FUNCTION_BLOCK EEE_Bruto (* Elevatoria de esgoto bruto - HidrycoLib *)
  (* Standard: 61499-2 *)
  (* Version 1.9, 21/10/2026, Hidryco, Hidryco, 1.9: Necessidade recebe o nivel em % (STS_NIVEL) para o grafico das faixas. 1.8: PID de nivel e velocidades da IHM/SCADA em Hz (conversao no CLP). 1.7: faixas da Necessidade e PID de nivel em % da altura do poco (LIT_100_03.stsPorcentagem). 1.6: pidCtl PidNivel com CycleTime 1000 ms (sem ele o calculo ciclico do pidSC ficava sem periodo). 1.5: variaveis de controle nos sub-CATs Necessidade, Revezamento e PID (padrao ElevatoriaEsgotoBruto); reset cmdResetFalhas / E_RESET_FALHAS_PROCESSO; PT_100_01, LSL_100_04, LSH_100_05 e pidCtl PidNivel. 1.4: simbolos sBoiaL/sBoiaH (boias animadas, verde/vermelho); velocidades na IHM em Hz. 1.3: selecao do gerador bomba por bomba (geradorHabilitaBS01/02/03, cada uma so na sua bomba; antes geradorHabilita unica). 1.2: emergencia do PCM NF (stsEmergenciaPainel FALSE = em emergencia, so depois da 1a leitura); FALHA UCP das bombas NF (cfgTermicaNF TRUE: FALSE no campo = falha); rede do CAT reorganizada. 1.1: emergencia do PCM pelo symlink ${PATH}stsEmergenciaPainel (soma com stsEmergencia do processo); comunicacao dos ATV630 pelos symlinks ${PATH}atvComunicacaoBS01..03 (ComStatus do HW CAT ATVSpeedControlMbtcp) publicada como ${PATH}BS_100_0x.stsFalhaComunicacao; cfgUsaFalhaComunicacao TRUE; estado 7 = emergencia. 1.0: elevatoria de esgoto bruto (3 bombas 100-BS-01/02/03, 2 + 1 reserva). Faixas de nivel do LIT-03, revezamento por tempo, velocidade pelo PID de nivel, HH do Nereda segura o esgoto ate o H do poco, operacao pelas boias com o LIT-03 em falha, falha de recalque pelo PIT-01. Campo por symlink ${PATH}: stsBoiaNivelBaixo (LSL-04), stsBoiaNivelAlto (LSH-05); bombas e sensores pelos symlinks dos proprios CATs (${PATH}BS_100_0x., ${PATH}LIT_100_03., ${PATH}PIT_100_01.). *)
  PACKAGE Hidryco.HidrycoLib;
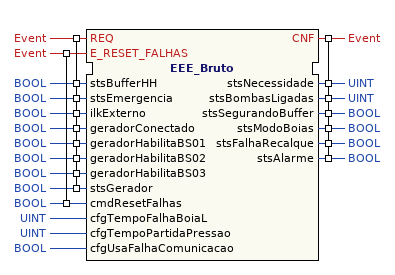
  EVENT_INPUT
    REQ WITH stsBufferHH, stsEmergencia, ilkExterno, geradorConectado, geradorHabilitaBS01, geradorHabilitaBS02, geradorHabilitaBS03, stsGerador; (* Atualizacao do processo *)
    E_RESET_FALHAS WITH cmdResetFalhas; (* Reset pelo processo (elevatoria, bombas e sensores) com cmdResetFalhas = TRUE *)
  END_EVENT
  EVENT_OUTPUT
    CNF WITH stsNecessidade, stsBombasLigadas, stsSegurandoBuffer, stsModoBoias, stsFalhaRecalque, stsAlarme; (* Status (so na mudanca) *)
  END_EVENT
  VAR_INPUT
    stsBufferHH : BOOL; (* Alarme HH do nivel do tanque de equalizacao do Nereda (40-LT-0001): a elevatoria segura o esgoto *)
    stsEmergencia : BOOL; (* Emergencia pelo processo (soma com a emergencia do PCM lida pelo symlink stsEmergenciaPainel): retira o comando das bombas *)
    ilkExterno : BOOL; (* Intertravamento externo do automatico das bombas (ex.: falha das UCTs, futuro) *)
    geradorConectado : BOOL; (* O gerador pode alimentar as bombas *)
    geradorHabilitaBS01 : BOOL; (* Bomba 100-BS-01 liberada para operar com a planta no gerador (HAB_BS_100_01 do CAT Subestacao) *)
    geradorHabilitaBS02 : BOOL; (* Bomba 100-BS-02 liberada para operar com a planta no gerador (HAB_BS_100_02 do CAT Subestacao) *)
    geradorHabilitaBS03 : BOOL; (* Bomba 100-BS-03 liberada para operar com a planta no gerador (HAB_BS_100_03 do CAT Subestacao) *)
    stsGerador : BOOL; (* Planta alimentada pelo gerador *)
    cmdResetFalhas : BOOL; (* TRUE = reset (com o evento E_RESET_FALHAS) *)
    cfgTempoFalhaBoiaL : UINT := 10; (* Operacao pelas boias com a boia LSL com defeito: bombas ficam ligadas este tempo (min) depois que a LSH desce *)
    cfgTempoPartidaPressao : UINT := 30; (* Alarmes L/LL do PIT-01 inibidos ate a bomba estar ligada ha este tempo (s); tambem inibidos com as bombas paradas *)
    cfgUsaFalhaComunicacao : BOOL := TRUE; (* Bombas: TRUE = falha de comunicacao com o ATV630 (symlink atvComunicacaoBS0x = ComStatus do HW CAT) tira a bomba do automatico *)
  END_VAR
  VAR_OUTPUT
    stsNecessidade : UINT; (* Numero de bombas pedidas (0, 1, 2) *)
    stsBombasLigadas : UINT; (* Bombas ligadas *)
    stsSegurandoBuffer : BOOL; (* Elevatoria parada segurando o esgoto (HH do tanque do Nereda) *)
    stsModoBoias : BOOL; (* Operacao de emergencia pelas boias (LIT-03 em falha) *)
    stsFalhaRecalque : BOOL; (* Falha de recalque (pressao LL com bomba ligada) - memorizada ate o reset *)
    stsAlarme : BOOL; (* Algum alarme da elevatoria *)
  END_VAR
  FBS
    IThis : EEE_Bruto_HMI(QI := TRUE);
    plcStart1 : plcStart(Prio := 10);
    Logica : basicEEEBruto;
    Tick : E_CYCLE(DT := T#1s);
    PidNivel : pidCtl(CycleTime := 1000, Direction := FALSE, Bump := FALSE, ProhibitOutInc := FALSE, ProhibitOutDec := FALSE);
    LIT_100_03 : Sensor_Generico(pin_FC98F78ABCBC0A7E := TRUE, pin_CC8EEC06FF0C4430 := 'm');
    PT_100_01 : Sensor_Generico(pin_CC8EEC06FF0C4430 := 'bar');
    LSL_100_04 : SYMLINKMULTIVARDST_1559B0FF8170C9BA0(NAME1 := '$${PATH}stsBoiaNivelBaixo', QI := TRUE); {SET_ATTRIBUTE(Configuration.GenericFBType.InterfaceParams, Runtime.System#I:=1;VALUE${I$}:BOOL)}
    LSH_100_05 : SYMLINKMULTIVARDST_1559B0FF8170C9BA0(NAME1 := '$${PATH}stsBoiaNivelAlto', QI := TRUE); {SET_ATTRIBUTE(Configuration.GenericFBType.InterfaceParams, Runtime.System#I:=1;VALUE${I$}:BOOL)}
    EmergenciaPainel : SYMLINKMULTIVARDST_1559B0FF8170C9BA0(NAME1 := '$${PATH}stsEmergenciaPainel', QI := TRUE); {SET_ATTRIBUTE(Configuration.GenericFBType.InterfaceParams, Runtime.System#I:=1;VALUE${I$}:BOOL)}
    BS_100_01 : Motor_Generico(pin_63EFEFB7C85EC93E := TRUE, pin_66763E13F70A4420 := TRUE, pin_D34C88BE7FFF3208 := TRUE, pin_1ECF468387CA7EB2 := 0.0, pin_540BE0E4E6611ACA := 100.0, pin_E24313AE3BEE4D49 := 0.0, pin_39489193B7758574 := 600.0);
    BS_100_02 : Motor_Generico(pin_63EFEFB7C85EC93E := TRUE, pin_66763E13F70A4420 := TRUE, pin_D34C88BE7FFF3208 := TRUE, pin_1ECF468387CA7EB2 := 0.0, pin_540BE0E4E6611ACA := 100.0, pin_E24313AE3BEE4D49 := 0.0, pin_39489193B7758574 := 600.0);
    BS_100_03 : Motor_Generico(pin_63EFEFB7C85EC93E := TRUE, pin_66763E13F70A4420 := TRUE, pin_D34C88BE7FFF3208 := TRUE, pin_1ECF468387CA7EB2 := 0.0, pin_540BE0E4E6611ACA := 100.0, pin_E24313AE3BEE4D49 := 0.0, pin_39489193B7758574 := 600.0);
    AlarmeRecalque : ALARM_BIT(TYPE := 1, ACKTYPE_1 := 2, ACTIVE := TRUE); {SET_ATTRIBUTE(HMI.AlarmText, Falha de recalque: pressão muito baixa com bomba ligada)}
    AlarmeNivelAlto : ALARM_BIT(TYPE := 1, ACKTYPE_1 := 2, ACTIVE := TRUE); {SET_ATTRIBUTE(HMI.AlarmText, Nível alto no poço (boia LSH))}
    AlarmeFalhaBoia : ALARM_BIT(TYPE := 1, ACKTYPE_1 := 2, ACTIVE := TRUE); {SET_ATTRIBUTE(HMI.AlarmText, Defeito na boia de nível baixo (LSL))} {SET_ATTRIBUTE(HMI.AlarmClass, Warning)}
    Necessidade : Controle_Necessidade;
    Revezamento : Controle_Revezamento_3;
    PID : Controle_PID;
  END_FBS
  EVENT_CONNECTIONS
    plcStart1.FIRST_INIT TO IThis.9E38A1961DA6B101;
    plcStart1.REDO_INIT TO IThis.9E38A1961DA6B101;
    IThis.5F0B40587FEFE3C8 TO Logica.2004138DB0750D97;
    Logica.5A945D0C0194930B TO Tick.START;
    Logica.5A945D0C0194930B TO LSL_100_04.INIT;
    Logica.5A945D0C0194930B TO LSH_100_05.INIT;
    Logica.5A945D0C0194930B TO EmergenciaPainel.INIT;
    Logica.5A945D0C0194930B TO AlarmeRecalque.INIT;
    AlarmeRecalque.INITO TO AlarmeRecalque.REQ_INITDATA;
    AlarmeRecalque.CNF_INITDATA TO AlarmeRecalque.ACTIVATE;
    AlarmeRecalque.INITO TO AlarmeNivelAlto.INIT;
    AlarmeNivelAlto.INITO TO AlarmeNivelAlto.REQ_INITDATA;
    AlarmeNivelAlto.CNF_INITDATA TO AlarmeNivelAlto.ACTIVATE;
    AlarmeNivelAlto.INITO TO AlarmeFalhaBoia.INIT;
    AlarmeFalhaBoia.INITO TO AlarmeFalhaBoia.REQ_INITDATA;
    AlarmeFalhaBoia.CNF_INITDATA TO AlarmeFalhaBoia.ACTIVATE;
    AlarmeFalhaBoia.INITO TO plcStart1.ACK_FIRST;
    IThis.6B160DD0F34FB9C9 TO Logica.42B63FD756FD5680;
    E_RESET_FALHAS TO Logica.7EBC1FDE51BD3B7B;
    E_RESET_FALHAS TO LIT_100_03.D21DAA5004F58516;
    E_RESET_FALHAS TO PT_100_01.D21DAA5004F58516;
    REQ TO Logica.0276E9EA951C8BF6;
    LIT_100_03.28A380156DB271B8 TO Logica.90222814CB973B20;
    LIT_100_03.28A380156DB271B8 TO PidNivel.REQ;
    PT_100_01.28A380156DB271B8 TO Logica.DBE1B2FFC7FF3B08;
    LSL_100_04.CNF TO Logica.6AC38C72D7780ED9;
    LSH_100_05.CNF TO Logica.6AC38C72D7780ED9;
    Tick.EO TO Logica.32C03C0D3ECD7A45;
    Logica.FC3525374D7CA084 TO PidNivel.REQ;
    PidNivel.CNF TO Logica.9F042AA84E34F103;
    PidNivel.C_CNF TO Logica.9F042AA84E34F103;
    Logica.94BCFE033FAC1A7D TO PT_100_01.33AD1B5E06E89E39;
    EmergenciaPainel.CNF TO Logica.24497764F9E7DCEC;
    BS_100_03.9D4F26EE27EDF5B9 TO Logica.FA43CD3D3768B370;
    Logica.248D4310F5B0BB17 TO CNF;
    Logica.1098D8AD1579135E TO IThis.8A9BE89122F8493C;
    Logica.ABCC05CB716E560A TO BS_100_01.21070E4B73BFECDC;
    REQ TO BS_100_01.21070E4B73BFECDC;
    E_RESET_FALHAS TO BS_100_01.BA30A65ADDA4ECC3;
    BS_100_01.9D4F26EE27EDF5B9 TO Logica.50C8D5E107305241;
    Logica.ABCC05CB716E560A TO BS_100_02.21070E4B73BFECDC;
    REQ TO BS_100_02.21070E4B73BFECDC;
    E_RESET_FALHAS TO BS_100_02.BA30A65ADDA4ECC3;
    BS_100_02.9D4F26EE27EDF5B9 TO Logica.50C8D5E107305241;
    Logica.ABCC05CB716E560A TO BS_100_03.21070E4B73BFECDC;
    REQ TO BS_100_03.21070E4B73BFECDC;
    E_RESET_FALHAS TO BS_100_03.BA30A65ADDA4ECC3;
    BS_100_03.9D4F26EE27EDF5B9 TO Logica.50C8D5E107305241;
    Logica.13609D02FAABDEC3 TO AlarmeRecalque.REQ;
    Logica.13609D02FAABDEC3 TO AlarmeNivelAlto.REQ;
    Logica.13609D02FAABDEC3 TO AlarmeFalhaBoia.REQ;
    AlarmeRecalque.IND_1 TO IThis.8A9BE89122F8493C;
    AlarmeNivelAlto.IND_1 TO IThis.8A9BE89122F8493C;
    AlarmeFalhaBoia.IND_1 TO IThis.8A9BE89122F8493C;
    IThis.6B160DD0F34FB9C9 TO AlarmeRecalque.ACK_C1;
    IThis.6B160DD0F34FB9C9 TO AlarmeNivelAlto.ACK_C1;
    IThis.6B160DD0F34FB9C9 TO AlarmeFalhaBoia.ACK_C1;
    BS_100_02.9D4F26EE27EDF5B9 TO Logica.FA43CD3D3768B370;
    BS_100_01.9D4F26EE27EDF5B9 TO Logica.FA43CD3D3768B370;
    Necessidade.0F2BD63F330E2BDA TO Logica.FF091F8ADF8E7596;
    Revezamento.B06A49437DB43D50 TO Logica.FF091F8ADF8E7596;
    PID.75EB05A15DC6DC61 TO Logica.FF091F8ADF8E7596;
    PID.75EB05A15DC6DC61 TO PidNivel.REQ_PARA;
    PID.75EB05A15DC6DC61 TO PidNivel.REQ_SP;
    AlarmeFalhaBoia.INITO TO Necessidade.BF5A5000C611AF6E;
    AlarmeFalhaBoia.INITO TO Revezamento.3E2B631069BF22E6;
    AlarmeFalhaBoia.INITO TO PID.117942CC3F34C94C;
    Logica.1098D8AD1579135E TO Necessidade.3304F06E342FF911;
    Logica.1098D8AD1579135E TO Revezamento.A7EEDA91D01D2772;
    Logica.1098D8AD1579135E TO PID.7BD84B0FC1882775;
  END_CONNECTIONS
  DATA_CONNECTIONS
    cfgTempoFalhaBoiaL TO Logica.2A75047CBF417CA4;
    cfgTempoPartidaPressao TO Logica.C074396BDF300B13;
    cmdResetFalhas TO Logica.2FA4CF278B4F3CB3;
    stsBufferHH TO Logica.63AE38B1858D4CE6;
    stsEmergencia TO Logica.36DCE701EB12A3D1;
    cmdResetFalhas TO LIT_100_03.1908F43CB878F5E7;
    cmdResetFalhas TO PT_100_01.1908F43CB878F5E7;
    LIT_100_03.D7422D307E6AF52D TO Logica.67419F14E8ECCCB2;
    LIT_100_03.726640D1704B3F86 TO Logica.52C92FD7A4E5C1FD;
    LIT_100_03.613F6EF6FA647237 TO Logica.D4A7159E837D53E2;
    PT_100_01.53279A5859ECAB18 TO Logica.6EC73A6F5DB8968E;
    Logica.C04015C0646E521D TO PT_100_01.A5CADABB487002E6;
    LSL_100_04.VALUE1 TO Logica.4A528109D2D85E74;
    LSH_100_05.VALUE1 TO Logica.0BE8A559782EECAE;
    EmergenciaPainel.VALUE1 TO Logica.994B7ED99B6C59BF;
    BS_100_01.0F3C10FA447A4A49 TO Logica.22DA8E3A7DE48F1A;
    BS_100_02.0F3C10FA447A4A49 TO Logica.EFA423F4EA5F0E53;
    BS_100_03.0F3C10FA447A4A49 TO Logica.E65C8A6E4484BF72;
    Logica.11F225DEC1D0B3A7 TO PidNivel.Mode;
    Logica.6DE3EFF6B05010A8 TO PidNivel.PresetValue;
    PidNivel.Out TO Logica.B9FF3BEF62466996;
    Logica.1F92935144C9F81B TO BS_100_01.87DAE15414E7C412;
    Logica.DB7819F9C5AF6F0F TO BS_100_01.F94ABA993E8E9FF4;
    Logica.51E32EDEA2ACC722 TO BS_100_01.8E1E39034B916602;
    ilkExterno TO BS_100_01.B35265D6C3CF40DC;
    Logica.F44BFB101D284D4B TO BS_100_01.85953C7B9294A9BF;
    geradorConectado TO BS_100_01.8914049066EE23D9;
    geradorHabilitaBS01 TO BS_100_01.5C3D51A654AD25BA;
    stsGerador TO BS_100_01.A33BC24B3E7310B0;
    cmdResetFalhas TO BS_100_01.C2F1E9C0FB076F17;
    cfgUsaFalhaComunicacao TO BS_100_01.3AD811F03C7B9855;
    BS_100_01.EBDC9E59C4286586 TO Logica.515A40650D020437;
    BS_100_01.40A5976BFB296133 TO Logica.466542BF0436C757;
    Logica.F7CBB0C674366AC9 TO BS_100_02.87DAE15414E7C412;
    Logica.DB7819F9C5AF6F0F TO BS_100_02.F94ABA993E8E9FF4;
    Logica.51E32EDEA2ACC722 TO BS_100_02.8E1E39034B916602;
    ilkExterno TO BS_100_02.B35265D6C3CF40DC;
    Logica.F44BFB101D284D4B TO BS_100_02.85953C7B9294A9BF;
    geradorConectado TO BS_100_02.8914049066EE23D9;
    geradorHabilitaBS02 TO BS_100_02.5C3D51A654AD25BA;
    stsGerador TO BS_100_02.A33BC24B3E7310B0;
    cmdResetFalhas TO BS_100_02.C2F1E9C0FB076F17;
    cfgUsaFalhaComunicacao TO BS_100_02.3AD811F03C7B9855;
    BS_100_02.EBDC9E59C4286586 TO Logica.AF1EF9EE1167DEDC;
    BS_100_02.40A5976BFB296133 TO Logica.FCA2071868470917;
    Logica.73409D95B7083780 TO BS_100_03.87DAE15414E7C412;
    Logica.DB7819F9C5AF6F0F TO BS_100_03.F94ABA993E8E9FF4;
    Logica.51E32EDEA2ACC722 TO BS_100_03.8E1E39034B916602;
    ilkExterno TO BS_100_03.B35265D6C3CF40DC;
    Logica.F44BFB101D284D4B TO BS_100_03.85953C7B9294A9BF;
    geradorConectado TO BS_100_03.8914049066EE23D9;
    geradorHabilitaBS03 TO BS_100_03.5C3D51A654AD25BA;
    stsGerador TO BS_100_03.A33BC24B3E7310B0;
    cmdResetFalhas TO BS_100_03.C2F1E9C0FB076F17;
    cfgUsaFalhaComunicacao TO BS_100_03.3AD811F03C7B9855;
    BS_100_03.EBDC9E59C4286586 TO Logica.5396A772225DEB3F;
    BS_100_03.40A5976BFB296133 TO Logica.9B8834E2710E7927;
    IThis.8DA339BF859A8E5F TO Logica.ECEAE676A6E41F28;
    Logica.AC7B9F1FA27C1FD1 TO AlarmeRecalque.INP;
    Logica.058FFE0E7D12B412 TO AlarmeNivelAlto.INP;
    Logica.3EF67A9DCF2789DB TO AlarmeFalhaBoia.INP;
    Logica.4AC7770F4C446AEA TO stsNecessidade;
    Logica.35666A9BF30FDCC7 TO stsBombasLigadas;
    Logica.E9F77451534DAE6C TO stsSegurandoBuffer;
    Logica.BF1AEE1747D48627 TO stsModoBoias;
    Logica.8F72D4456BAA5444 TO stsFalhaRecalque;
    Logica.E964EB18E69985AA TO stsAlarme;
    Logica.C9E401CFFAA6182F TO IThis.850B1619B9DA198C;
    Logica.A03F17C59577EA19 TO IThis.944B5897BE0574B9;
    Logica.35666A9BF30FDCC7 TO IThis.2C1A9CF4B602EE39;
    Logica.A676EAE8813C9472 TO IThis.7E6F53D9C30EBF39;
    Logica.93034EF747C7C8B2 TO IThis.65049BBD5A4BB493;
    Logica.BF1AEE1747D48627 TO IThis.AF62408DEC77723C;
    Logica.E9F77451534DAE6C TO IThis.291D653F26E2F3DA;
    Logica.8F72D4456BAA5444 TO IThis.61AA8C54482A7A9B;
    Logica.417E0C30BAF102DF TO IThis.EE7C6C6858FFBB22;
    Logica.173E069DE197A4CF TO IThis.AAD965D400369960;
    Logica.489475EDA9AC9EE5 TO IThis.FE4CB77CC09B077D;
    Logica.1ADD872C67BB4DE1 TO IThis.AFD72C4363D47798;
    Logica.13FC107471B9CC29 TO IThis.23E5A2CBCEA0A47D;
    Logica.E964EB18E69985AA TO IThis.55636688498925A1;
    AlarmeRecalque.STATE_1 TO IThis.8C8C7B22E6752219;
    AlarmeNivelAlto.STATE_1 TO IThis.458D5DB98E9425A3;
    AlarmeFalhaBoia.STATE_1 TO IThis.0DFF34EDE3D642CE;
    PID.C9DF845DD1ECA932 TO PidNivel.Sp;
    PID.4F45CBCE24FA8775 TO PidNivel.Gain;
    PID.5D86C7647B367BF7 TO PidNivel.IntegralTime;
    PID.C753842CF6C65D61 TO PidNivel.DerivativeTime;
    PID.8B11A5B11AA557C3 TO PidNivel.OutMin;
    PID.8B11A5B11AA557C3 TO Logica.39D99F13A06DDE55;
    PID.E7AF90225A9267BD TO PidNivel.OutMax;
    PID.E7AF90225A9267BD TO Logica.6FE815DDF49B081F;
    PID.004F03C1536C2B1E TO Logica.9E10D0E429B4004A;
    Necessidade.F8E4EB0276D578DB TO Logica.C05E87D9971F8886;
    Necessidade.5126CE4A870E517F TO Logica.8EB441F793280592;
    Necessidade.FCED367007BA1689 TO Logica.072A6C97AFD6585F;
    Necessidade.4B45B05E6464EEE7 TO Logica.BEFB8DAF08C8995F;
    Necessidade.B1260102A6291D33 TO Logica.7DBB130FE6E6C808;
    Revezamento.14B34C1C3DE79269 TO Logica.5A7C86072FF3CD5A;
    Revezamento.E9B6E434B3B859BA TO Logica.CCF7F3F47A1A1320;
    Revezamento.5B68F5BBF5994362 TO Logica.665448845ED3554E;
    Revezamento.49A70042A34A21C7 TO Logica.06814213D61A9713;
    Revezamento.1EA41783712558AD TO Logica.54CD99170D68F8C4;
    Logica.4AC7770F4C446AEA TO Necessidade.26BC67DB3AB94B29;
    Logica.172630242E663B7D TO Revezamento.7A2503B7B1388DC6;
    Logica.7CE98D61C5896B6B TO Revezamento.D93AFAFEC8E31E85;
    Logica.FB21944AFA623D56 TO Revezamento.E430C3F15AEF6E1E;
    Logica.02A0E42D87C41BFD TO PID.260D6E81A1639D84;
    LIT_100_03.E6F78A591442B69F TO Logica.0E2F0D9F0929276A;
    LIT_100_03.E6F78A591442B69F TO PidNivel.Pv;
    Logica.FEB697ACC839FDA4 TO IThis.51564348690894F5;
    LIT_100_03.E6F78A591442B69F TO Necessidade.26C50C1A131DC8B6;
  END_CONNECTIONS
END_FUNCTION_BLOCK
